(* IEC 61131-3 sources: codesys-api/examples/codesys4/projects/feature_probe.fbsdev/Application.iecapp^, 2 files *)

(* ---- PRG_Comms.prg.st ---- *)
PROGRAM PRG_Comms
VAR
    tcpClient : ModbusFB.ClientTCP;
    serialClient : ModbusFB.ClientSerial;
    readHolding : ModbusFB.ClientRequestReadHoldingRegisters;
    registers : ARRAY[0..9] OF UINT;
    comHandle : SysCom.RTS_IEC_HANDLE;
    comResult : SysCom.RTS_IEC_RESULT;
    mqttClient : MQTT.MQTTClient;
    jsonWriter : JSON.JSONByteArrayWriter;
    serverIp : ARRAY[0..3] OF BYTE := [192, 168, 50, 10];
END_VAR
tcpClient(xConnect := TRUE, aIPAddr := serverIp, uiPort := 502);
readHolding(rClient := tcpClient, uiUnitId := 1, uiStartItem := 0, uiQuantity := 10,
    pData := ADR(registers), xExecute := TRUE);
END_PROGRAM

(* ---- PRG_Control.prg.st ---- *)
PROGRAM PRG_Control
VAR RETAIN
    retainedCount : UDINT;
END_VAR
VAR PERSISTENT
    lastCommandId : UDINT;
END_VAR
VAR
    nowMs : UDINT;
    timestamp : ULINT;
    rtcResult : UDINT;
    dynamicBuffer : POINTER TO BYTE;
END_VAR
retainedCount := retainedCount + 1;
nowMs := SysTimeCore.SysTimeGetMs();
rtcResult := SysTimeRtc.SysTimeRtcHighResGet(pTimestamp := timestamp);
lastCommandId := lastCommandId + 1;
END_PROGRAM
